DATA_BLOCK "Main_DB"
{ S7_Optimized_Access := 'TRUE' }
VERSION : 0.1
"Main"

BEGIN

END_DATA_BLOCK
